Staubli VAL3: start.pgx

program start()
begin
  userPage("InOut")
end
